// TIA Portal V21 export
// export: Created 2026-05-12T00:00:00.0000000Z, ExportSetting None
DATA_BLOCK "DB_HMI_Interface"   // DB200
TITLE = DB title
{ S7_Optimized_Access := 'FALSE' }
// 保持注释
   VAR
      Enabled : Bool := false;
   END_VAR
   VAR RETAIN
      DefaultInt : Int;   // Retained setpoint / 保持设定值
   END_VAR
   VAR
      "电机/运行%2F" : Bool := true;
      Motor : Struct
         Config : Struct
            Speed : Real := 1.5;
         END_STRUCT;
      END_STRUCT;
      Samples : Array[0..1] of Int;
      Locked : Int := 7;
      Inherited : Struct
         Value : Int;
      END_STRUCT;
      LockedValue : Int := 9;
      Typed : "MotorType";
      Clock : DTL;
      ConstantLiteral : Int := 42;
      BulkValue : Int := 2(4);
      Hardware : HW_IO := 64;
      AnyDb : DB_ANY := 42;
      SymbolicText : String[MaxText] := 'alpha';
      HardwareExpression : HW_IO := ModuleName;
      DefaultHardware : HW_IO;
   END_VAR
BEGIN
   Samples[0] := 3;
   Typed.NestedValue := 5;
END_DATA_BLOCK
